Staubli VAL3: deleteItem.pgx

public program deleteItem()
  local string l_sMsg
  local bool l_bResult
begin
  if sSelTraj!=""
    l_sMsg="是否删除："+sSelTraj+"?"
    l_bResult=userPageConfirm(l_sMsg)
    if l_bResult
      call trajectory:deleteTraj(sSelTraj,bToSave)
      //call trajectory:getTrajList(sList)
    endIf
  else
    userPageAlert("未选中任意项目！")
  endIf
end
